{attribute 'pack_mode' := '1'}
TYPE ST_MqttCommand_Rx :
STRUCT	// 인터페이스 100.Command 버전 2 (2026-11-25): 16 B, SequenceNumber 없음
	DeviceIndex	:	UDINT;	// 장치 번호 1부터 (F_MqttDistribute가 레코드 맨 앞에서 읽음: nIndexOffset = 0)
	CommandType	:	UDINT;
	Value		:	REAL;	// kW 등, CommandType에 따라 의미가 다름
	Delay		:	UDINT;	// ms. 이만큼 기다렸다가 실행 (0이면 바로). FB_EmsCmdGate
END_STRUCT
END_TYPE

(* stored: Version 1.1.0.1, ProductVersion 3.1.4024.9
   DUT ST_MqttCommand_Rx: Id {151a57c0-4a25-41d6-bd3b-a15635e8751f} *)
